  movel([-0.151447, -0.828061, -2.797798, -1.086530, 1.570796, 1.419350],accel_mss,speed_ms,0,blend_radius_m)
  movel([-0.155435, -0.836303, -2.796291, -1.079795, 1.570796, 1.415362],accel_mss,speed_ms,0,blend_radius_m)
  movel([-0.157149, -0.840333, -2.795540, -1.076516, 1.570796, 1.413648],accel_mss,speed_ms,0,blend_radius_m)
  movel([-0.159989, -0.848193, -2.794051, -1.070145, 1.570796, 1.410807],accel_mss,speed_ms,0,blend_radius_m)
  movel([-0.161109, -0.852028, -2.793312, -1.067049, 1.570796, 1.409688],accel_mss,speed_ms,0,blend_radius_m)
  movel([-0.162732, -0.859501, -2.791847, -1.061041, 1.570796, 1.408064],accel_mss,speed_ms,0,blend_radius_m)
  movel([-0.163230, -0.863145, -2.791122, -1.058122, 1.570796, 1.407566],accel_mss,speed_ms,0,blend_radius_m)
  movel([-0.163513, -0.866720, -2.790402, -1.055267, 1.570796, 1.407283],accel_mss,speed_ms,0,blend_radius_m)
  movel([-0.163602, -0.871655, -2.789397, -1.051337, 1.570796, 1.407194],accel_mss,speed_ms,0,blend_radius_m)
  movel([-0.163380, -0.876401, -2.788417, -1.047571, 1.570796, 1.407417],accel_mss,speed_ms,0,blend_radius_m)
  movel([-0.162870, -0.880943, -2.787467, -1.043979, 1.570796, 1.407926],accel_mss,speed_ms,0,blend_radius_m)
  movel([-0.162104, -0.885286, -2.786547, -1.040556, 1.570796, 1.408692],accel_mss,speed_ms,0,blend_radius_m)
  movel([-0.161097, -0.889404, -2.785664, -1.037321, 1.570796, 1.409700],accel_mss,speed_ms,0,blend_radius_m)
  movel([-0.159870, -0.893285, -2.784823, -1.034282, 1.570796, 1.410927],accel_mss,speed_ms,0,blend_radius_m)
  movel([-0.158448, -0.896924, -2.784025, -1.031439, 1.570796, 1.412348],accel_mss,speed_ms,0,blend_radius_m)
  movel([-0.156848, -0.900304, -2.783277, -1.028807, 1.570796, 1.413948],accel_mss,speed_ms,0,blend_radius_m)
  movel([-0.149158, -0.912135, -2.780604, -1.019650, 1.570796, 1.421638],accel_mss,speed_ms,0,blend_radius_m)
  movel([-0.143209, -0.921779, -2.778359, -1.012250, 1.570796, 1.427587],accel_mss,speed_ms,0,blend_radius_m)
  movel([-0.142775, -0.922813, -2.778115, -1.011461, 1.570796, 1.428021],accel_mss,speed_ms,0,blend_radius_m)
  movel([-0.135600, -0.913354, -2.780324, -1.018712, 1.570796, 1.435197],accel_mss,speed_ms,0,blend_radius_m)
  movel([-0.127938, -0.904013, -2.782449, -1.025928, 1.570796, 1.442859],accel_mss,speed_ms,0,blend_radius_m)
  movel([-0.119839, -0.894825, -2.784486, -1.033078, 1.570796, 1.450957],accel_mss,speed_ms,0,blend_radius_m)
  movel([-0.111369, -0.885835, -2.786430, -1.040124, 1.570796, 1.459427],accel_mss,speed_ms,0,blend_radius_m)
  movel([-0.102591, -0.877095, -2.788273, -1.047021, 1.570796, 1.468205],accel_mss,speed_ms,0,blend_radius_m)
  movel([-0.093574, -0.868644, -2.790012, -1.053733, 1.570796, 1.477222],accel_mss,speed_ms,0,blend_radius_m)
  movel([-0.084386, -0.860539, -2.791641, -1.060208, 1.570796, 1.486410],accel_mss,speed_ms,0,blend_radius_m)
  movel([-0.075105, -0.852829, -2.793156, -1.066404, 1.570796, 1.495692],accel_mss,speed_ms,0,blend_radius_m)
  movel([-0.070692, -0.849394, -2.793820, -1.069175, 1.570796, 1.500104],accel_mss,speed_ms,0,blend_radius_m)
  movel([-0.066171, -0.846121, -2.794447, -1.071821, 1.570796, 1.504626],accel_mss,speed_ms,0,blend_radius_m)
  movel([-0.061579, -0.843047, -2.795030, -1.074312, 1.570796, 1.509218],accel_mss,speed_ms,0,blend_radius_m)
  movel([-0.056967, -0.840218, -2.795562, -1.076609, 1.570796, 1.513830],accel_mss,speed_ms,0,blend_radius_m)
  movel([-0.052375, -0.837673, -2.796037, -1.078679, 1.570796, 1.518421],accel_mss,speed_ms,0,blend_radius_m)
  movel([-0.047846, -0.835454, -2.796448, -1.080487, 1.570796, 1.522951],accel_mss,speed_ms,0,blend_radius_m)
  movel([-0.043425, -0.833599, -2.796789, -1.082000, 1.570796, 1.527371],accel_mss,speed_ms,0,blend_radius_m)
  movel([-0.039161, -0.832150, -2.797055, -1.083184, 1.570796, 1.531636],accel_mss,speed_ms,0,blend_radius_m)
  movel([-0.035094, -0.831147, -2.797238, -1.084004, 1.570796, 1.535702],accel_mss,speed_ms,0,blend_radius_m)
  movel([-0.031268, -0.830626, -2.797333, -1.084430, 1.570796, 1.539528],accel_mss,speed_ms,0,blend_radius_m)
  movel([-0.027734, -0.830629, -2.797332, -1.084428, 1.570796, 1.543062],accel_mss,speed_ms,0,blend_radius_m)
  movel([-0.024533, -0.831189, -2.797230, -1.083970, 1.570796, 1.546264],accel_mss,speed_ms,0,blend_radius_m)
  movel([-0.021709, -0.832340, -2.797020, -1.083029, 1.570796, 1.549087],accel_mss,speed_ms,0,blend_radius_m)
  movel([-0.019297, -0.834113, -2.796695, -1.081581, 1.570796, 1.551499],accel_mss,speed_ms,0,blend_radius_m)
  movel([-0.017345, -0.836537, -2.796247, -1.079604, 1.570796, 1.553452],accel_mss,speed_ms,0,blend_radius_m)
  movel([-0.015891, -0.839644, -2.795669, -1.077075, 1.570796, 1.554905],accel_mss,speed_ms,0,blend_radius_m)
  movel([-0.014708, -0.844472, -2.794760, -1.073157, 1.570796, 1.556088],accel_mss,speed_ms,0,blend_radius_m)
  movel([-0.014174, -0.849958, -2.793712, -1.068720, 1.570796, 1.556622],accel_mss,speed_ms,0,blend_radius_m)
  movel([-0.014196, -0.855947, -2.792548, -1.063895, 1.570796, 1.556600],accel_mss,speed_ms,0,blend_radius_m)
  movel([-0.014673, -0.862293, -2.791292, -1.058804, 1.570796, 1.556123],accel_mss,speed_ms,0,blend_radius_m)
  movel([-0.015515, -0.868851, -2.789970, -1.053568, 1.570796, 1.555282],accel_mss,speed_ms,0,blend_radius_m)
  movel([-0.016634, -0.875486, -2.788607, -1.048296, 1.570796, 1.554162],accel_mss,speed_ms,0,blend_radius_m)
  movel([-0.019330, -0.888444, -2.785871, -1.038074, 1.570796, 1.551466],accel_mss,speed_ms,0,blend_radius_m)
  movel([-0.021385, -0.896660, -2.784083, -1.031646, 1.570796, 1.549411],accel_mss,speed_ms,0,blend_radius_m)
  movel([-0.023782, -0.904827, -2.782265, -1.025296, 1.570796, 1.547015],accel_mss,speed_ms,0,blend_radius_m)
  movel([-0.026474, -0.912947, -2.780417, -1.019025, 1.570796, 1.544323],accel_mss,speed_ms,0,blend_radius_m)
  movel([-0.029419, -0.921037, -2.778534, -1.012818, 1.570796, 1.541377],accel_mss,speed_ms,0,blend_radius_m)
  movel([-0.032573, -0.929096, -2.776617, -1.006676, 1.570796, 1.538223],accel_mss,speed_ms,0,blend_radius_m)
  movel([-0.035892, -0.937137, -2.774661, -1.000590, 1.570796, 1.534904],accel_mss,speed_ms,0,blend_radius_m)
  movel([-0.042880, -0.953213, -2.770623, -0.988553, 1.570796, 1.527916],accel_mss,speed_ms,0,blend_radius_m)
  movel([-0.036325, -0.953508, -2.770548, -0.988333, 1.570796, 1.534471],accel_mss,speed_ms,0,blend_radius_m)
  movel([-0.032953, -0.953917, -2.770442, -0.988029, 1.570796, 1.537843],accel_mss,speed_ms,0,blend_radius_m)
  movel([-0.030089, -0.954829, -2.770208, -0.987352, 1.570796, 1.540707],accel_mss,speed_ms,0,blend_radius_m)
  movel([-0.028984, -0.955552, -2.770021, -0.986816, 1.570796, 1.541813],accel_mss,speed_ms,0,blend_radius_m)
  movel([-0.028168, -0.956495, -2.769777, -0.986117, 1.570796, 1.542628],accel_mss,speed_ms,0,blend_radius_m)
  movel([-0.027690, -0.957681, -2.769470, -0.985239, 1.570796, 1.543106],accel_mss,speed_ms,0,blend_radius_m)
  movel([-0.027603, -0.959140, -2.769090, -0.984159, 1.570796, 1.543193],accel_mss,speed_ms,0,blend_radius_m)
  movel([-0.027958, -0.960895, -2.768632, -0.982862, 1.570796, 1.542838],accel_mss,speed_ms,0,blend_radius_m)
  movel([-0.028810, -0.962986, -2.768083, -0.981321, 1.570796, 1.541986],accel_mss,speed_ms,0,blend_radius_m)
  movel([-0.030204, -0.965433, -2.767436, -0.979520, 1.570796, 1.540592],accel_mss,speed_ms,0,blend_radius_m)
  movel([-0.032189, -0.968258, -2.766684, -0.977447, 1.570796, 1.538607],accel_mss,speed_ms,0,blend_radius_m)
  movel([-0.034030, -0.970557, -2.766069, -0.975764, 1.570796, 1.536766],accel_mss,speed_ms,0,blend_radius_m)
  movel([-0.035882, -0.972625, -2.765511, -0.974253, 1.570796, 1.534914],accel_mss,speed_ms,0,blend_radius_m)
  movel([-0.037742, -0.974479, -2.765009, -0.972901, 1.570796, 1.533055],accel_mss,speed_ms,0,blend_radius_m)
  movel([-0.041487, -0.977625, -2.764152, -0.970612, 1.570796, 1.529310],accel_mss,speed_ms,0,blend_radius_m)
  movel([-0.043369, -0.978954, -2.763787, -0.969648, 1.570796, 1.527427],accel_mss,speed_ms,0,blend_radius_m)
  movel([-0.047159, -0.981220, -2.763163, -0.968006, 1.570796, 1.523638],accel_mss,speed_ms,0,blend_radius_m)
  movel([-0.050963, -0.983074, -2.762650, -0.966665, 1.570796, 1.519833],accel_mss,speed_ms,0,blend_radius_m)
  movel([-0.054779, -0.984659, -2.762209, -0.965521, 1.570796, 1.516017],accel_mss,speed_ms,0,blend_radius_m)
  movel([-0.062394, -0.987558, -2.761398, -0.963434, 1.570796, 1.508402],accel_mss,speed_ms,0,blend_radius_m)
  movel([-0.066370, -0.993967, -2.759582, -0.958840, 1.570796, 1.504426],accel_mss,speed_ms,0,blend_radius_m)
  movel([-0.068546, -0.997167, -2.758665, -0.956558, 1.570796, 1.502250],accel_mss,speed_ms,0,blend_radius_m)
  movel([-0.070857, -1.000276, -2.757766, -0.954347, 1.570796, 1.499939],accel_mss,speed_ms,0,blend_radius_m)
  movel([-0.073309, -1.003227, -2.756906, -0.952256, 1.570796, 1.497488],accel_mss,speed_ms,0,blend_radius_m)
  movel([-0.075903, -1.005952, -2.756106, -0.950331, 1.570796, 1.494894],accel_mss,speed_ms,0,blend_radius_m)
  movel([-0.078648, -1.008386, -2.755387, -0.948616, 1.570796, 1.492149],accel_mss,speed_ms,0,blend_radius_m)
  movel([-0.081555, -1.010470, -2.754767, -0.947152, 1.570796, 1.489241],accel_mss,speed_ms,0,blend_radius_m)
  movel([-0.083598, -1.011520, -2.754454, -0.946415, 1.570796, 1.487198],accel_mss,speed_ms,0,blend_radius_m)
  movel([-0.085214, -1.011878, -2.754347, -0.946164, 1.570796, 1.485582],accel_mss,speed_ms,0,blend_radius_m)
  movel([-0.086450, -1.011645, -2.754417, -0.946328, 1.570796, 1.484347],accel_mss,speed_ms,0,blend_radius_m)
  movel([-0.087346, -1.010917, -2.754634, -0.946838, 1.570796, 1.483451],accel_mss,speed_ms,0,blend_radius_m)
  movel([-0.087946, -1.009791, -2.754969, -0.947628, 1.570796, 1.482851],accel_mss,speed_ms,0,blend_radius_m)
  movel([-0.088287, -1.008371, -2.755391, -0.948627, 1.570796, 1.482509],accel_mss,speed_ms,0,blend_radius_m)
  movel([-0.088418, -1.006753, -2.755870, -0.949766, 1.570796, 1.482378],accel_mss,speed_ms,0,blend_radius_m)
  movel([-0.088369, -1.005030, -2.756377, -0.950982, 1.570796, 1.482428],accel_mss,speed_ms,0,blend_radius_m)
  movel([-0.087893, -1.001208, -2.757495, -0.953686, 1.570796, 1.482904],accel_mss,speed_ms,0,blend_radius_m)
  movel([-0.087059, -0.997250, -2.758641, -0.956499, 1.570796, 1.483737],accel_mss,speed_ms,0,blend_radius_m)
  movel([-0.084858, -0.988993, -2.760994, -0.962402, 1.570796, 1.485939],accel_mss,speed_ms,0,blend_radius_m)
  movel([-0.093540, -0.987568, -2.761395, -0.963426, 1.570796, 1.477256],accel_mss,speed_ms,0,blend_radius_m)
  movel([-0.102455, -0.986524, -2.761688, -0.964178, 1.570796, 1.468341],accel_mss,speed_ms,0,blend_radius_m)
  movel([-0.111365, -0.985448, -2.761989, -0.964952, 1.570796, 1.459431],accel_mss,speed_ms,0,blend_radius_m)
  movel([-0.115747, -0.984770, -2.762178, -0.965441, 1.570796, 1.455049],accel_mss,speed_ms,0,blend_radius_m)
  movel([-0.120046, -0.983927, -2.762413, -0.966049, 1.570796, 1.450750],accel_mss,speed_ms,0,blend_radius_m)
  movel([-0.124039, -0.982910, -2.762695, -0.966783, 1.570796, 1.446757],accel_mss,speed_ms,0,blend_radius_m)
  movel([-0.127889, -0.981713, -2.763027, -0.967649, 1.570796, 1.442907],accel_mss,speed_ms,0,blend_radius_m)
  movel([-0.135327, -0.978974, -2.763782, -0.969633, 1.570796, 1.435469],accel_mss,speed_ms,0,blend_radius_m)
  movel([-0.142709, -0.976168, -2.764550, -0.971671, 1.570796, 1.428087],accel_mss,speed_ms,0,blend_radius_m)
  movel([-0.150371, -0.973750, -2.765207, -0.973432, 1.570796, 1.420425],accel_mss,speed_ms,0,blend_radius_m)
  movel([-0.152086, -0.978530, -2.763904, -0.969955, 1.570796, 1.418710],accel_mss,speed_ms,0,blend_radius_m)
  movel([-0.153549, -0.983185, -2.762619, -0.966585, 1.570796, 1.417247],accel_mss,speed_ms,0,blend_radius_m)
  movel([-0.154762, -0.987705, -2.761356, -0.963328, 1.570796, 1.416035],accel_mss,speed_ms,0,blend_radius_m)
  movel([-0.155729, -0.992084, -2.760119, -0.960186, 1.570796, 1.415067],accel_mss,speed_ms,0,blend_radius_m)
  movel([-0.156451, -0.996319, -2.758909, -0.957161, 1.570796, 1.414345],accel_mss,speed_ms,0,blend_radius_m)
  movel([-0.156938, -1.000405, -2.757728, -0.954256, 1.570796, 1.413859],accel_mss,speed_ms,0,blend_radius_m)
  movel([-0.157185, -1.004336, -2.756581, -0.951472, 1.570796, 1.413612],accel_mss,speed_ms,0,blend_radius_m)
  movel([-0.157205, -1.008112, -2.755468, -0.948809, 1.570796, 1.413592],accel_mss,speed_ms,0,blend_radius_m)
  movel([-0.156995, -1.011726, -2.754393, -0.946271, 1.570796, 1.413802],accel_mss,speed_ms,0,blend_radius_m)
  movel([-0.156554, -1.015168, -2.753359, -0.943862, 1.570796, 1.414242],accel_mss,speed_ms,0,blend_radius_m)
  movel([-0.155895, -1.018445, -2.752366, -0.941578, 1.570796, 1.414901],accel_mss,speed_ms,0,blend_radius_m)
  movel([-0.155018, -1.021546, -2.751419, -0.939423, 1.570796, 1.415778],accel_mss,speed_ms,0,blend_radius_m)
  movel([-0.153919, -1.024464, -2.750522, -0.937404, 1.570796, 1.416877],accel_mss,speed_ms,0,blend_radius_m)
  movel([-0.152607, -1.027203, -2.749673, -0.935513, 1.570796, 1.418189],accel_mss,speed_ms,0,blend_radius_m)
  movel([-0.151084, -1.029753, -2.748877, -0.933759, 1.570796, 1.419713],accel_mss,speed_ms,0,blend_radius_m)
  movel([-0.149346, -1.032112, -2.748136, -0.932140, 1.570796, 1.421450],accel_mss,speed_ms,0,blend_radius_m)
  movel([-0.146282, -1.035378, -2.747104, -0.929908, 1.570796, 1.424514],accel_mss,speed_ms,0,blend_radius_m)
  movel([-0.142850, -1.038167, -2.746215, -0.928007, 1.570796, 1.427946],accel_mss,speed_ms,0,blend_radius_m)
  movel([-0.139097, -1.040532, -2.745456, -0.926400, 1.570796, 1.431699],accel_mss,speed_ms,0,blend_radius_m)
  movel([-0.135055, -1.042514, -2.744817, -0.925058, 1.570796, 1.435741],accel_mss,speed_ms,0,blend_radius_m)
  movel([-0.130770, -1.044161, -2.744284, -0.923944, 1.570796, 1.440026],accel_mss,speed_ms,0,blend_radius_m)
  movel([-0.126280, -1.045512, -2.743844, -0.923033, 1.570796, 1.444516],accel_mss,speed_ms,0,blend_radius_m)
  movel([-0.121626, -1.046612, -2.743485, -0.922291, 1.570796, 1.449171],accel_mss,speed_ms,0,blend_radius_m)
  movel([-0.116838, -1.047491, -2.743198, -0.921700, 1.570796, 1.453958],accel_mss,speed_ms,0,blend_radius_m)
  movel([-0.106974, -1.048821, -2.742762, -0.920806, 1.570796, 1.463822],accel_mss,speed_ms,0,blend_radius_m)
  movel([-0.096981, -1.049909, -2.742404, -0.920076, 1.570796, 1.473815],accel_mss,speed_ms,0,blend_radius_m)
  movel([-0.089406, -1.051010, -2.742041, -0.919338, 1.570796, 1.481391],accel_mss,speed_ms,0,blend_radius_m)
  movel([-0.086797, -1.051182, -2.741984, -0.919223, 1.570796, 1.484000],accel_mss,speed_ms,0,blend_radius_m)
  movel([-0.082087, -1.051090, -2.742014, -0.919284, 1.570796, 1.488709],accel_mss,speed_ms,0,blend_radius_m)
  movel([-0.081105, -1.051267, -2.741956, -0.919166, 1.570796, 1.489692],accel_mss,speed_ms,0,blend_radius_m)
  movel([-0.080223, -1.051641, -2.741832, -0.918916, 1.570796, 1.490574],accel_mss,speed_ms,0,blend_radius_m)
  movel([-0.079458, -1.052276, -2.741622, -0.918491, 1.570796, 1.491338],accel_mss,speed_ms,0,blend_radius_m)
  movel([-0.078830, -1.053233, -2.741305, -0.917851, 1.570796, 1.491966],accel_mss,speed_ms,0,blend_radius_m)
  movel([-0.078371, -1.054578, -2.740857, -0.916954, 1.570796, 1.492426],accel_mss,speed_ms,0,blend_radius_m)
  movel([-0.078211, -1.056102, -2.740348, -0.915938, 1.570796, 1.492585],accel_mss,speed_ms,0,blend_radius_m)
  movel([-0.078322, -1.057772, -2.739789, -0.914828, 1.570796, 1.492474],accel_mss,speed_ms,0,blend_radius_m)
  movel([-0.078680, -1.059571, -2.739183, -0.913635, 1.570796, 1.492116],accel_mss,speed_ms,0,blend_radius_m)
  movel([-0.079260, -1.061466, -2.738542, -0.912381, 1.570796, 1.491536],accel_mss,speed_ms,0,blend_radius_m)
  movel([-0.080989, -1.065467, -2.737179, -0.909743, 1.570796, 1.489808],accel_mss,speed_ms,0,blend_radius_m)
  movel([-0.082090, -1.067524, -2.736473, -0.908392, 1.570796, 1.488706],accel_mss,speed_ms,0,blend_radius_m)
  movel([-0.084632, -1.071630, -2.735052, -0.905706, 1.570796, 1.486165],accel_mss,speed_ms,0,blend_radius_m)
  movel([-0.087485, -1.075584, -2.733670, -0.903134, 1.570796, 1.483311],accel_mss,speed_ms,0,blend_radius_m)
  movel([-0.090454, -1.079207, -2.732393, -0.900789, 1.570796, 1.480342],accel_mss,speed_ms,0,blend_radius_m)
  movel([-0.093367, -1.082332, -2.731281, -0.898775, 1.570796, 1.477429],accel_mss,speed_ms,0,blend_radius_m)
  movel([-0.097927, -1.086556, -2.729766, -0.896068, 1.570796, 1.472870],accel_mss,speed_ms,0,blend_radius_m)
  movel([-0.100289, -1.088512, -2.729058, -0.894819, 1.570796, 1.470507],accel_mss,speed_ms,0,blend_radius_m)
  movel([-0.102689, -1.090353, -2.728389, -0.893647, 1.570796, 1.468107],accel_mss,speed_ms,0,blend_radius_m)
  movel([-0.107574, -1.093687, -2.727170, -0.891532, 1.570796, 1.463222],accel_mss,speed_ms,0,blend_radius_m)
  movel([-0.112504, -1.096527, -2.726124, -0.889738, 1.570796, 1.458292],accel_mss,speed_ms,0,blend_radius_m)
  movel([-0.117406, -1.098838, -2.725267, -0.888284, 1.570796, 1.453391],accel_mss,speed_ms,0,blend_radius_m)
  movel([-0.122195, -1.100585, -2.724616, -0.887188, 1.570796, 1.448602],accel_mss,speed_ms,0,blend_radius_m)
  movel([-0.124527, -1.101233, -2.724374, -0.886782, 1.570796, 1.446270],accel_mss,speed_ms,0,blend_radius_m)
  movel([-0.129018, -1.102060, -2.724064, -0.886265, 1.570796, 1.441778],accel_mss,speed_ms,0,blend_radius_m)
  movel([-0.131158, -1.102227, -2.724002, -0.886161, 1.570796, 1.439638],accel_mss,speed_ms,0,blend_radius_m)
  movel([-0.133875, -1.102203, -2.724010, -0.886175, 1.570796, 1.436921],accel_mss,speed_ms,0,blend_radius_m)
  movel([-0.136457, -1.101939, -2.724110, -0.886341, 1.570796, 1.434339],accel_mss,speed_ms,0,blend_radius_m)
  movel([-0.138916, -1.101462, -2.724288, -0.886639, 1.570796, 1.431880],accel_mss,speed_ms,0,blend_radius_m)
  movel([-0.141274, -1.100811, -2.724531, -0.887046, 1.570796, 1.429522],accel_mss,speed_ms,0,blend_radius_m)
  movel([-0.145748, -1.099110, -2.725166, -0.888114, 1.570796, 1.425048],accel_mss,speed_ms,0,blend_radius_m)
  movel([-0.150009, -1.097098, -2.725912, -0.889378, 1.570796, 1.420787],accel_mss,speed_ms,0,blend_radius_m)
  movel([-0.155186, -1.094353, -2.726925, -0.891111, 1.570796, 1.415610],accel_mss,speed_ms,0,blend_radius_m)
  movel([-0.160187, -1.091303, -2.728043, -0.893043, 1.570796, 1.410610],accel_mss,speed_ms,0,blend_radius_m)
  movel([-0.164967, -1.087926, -2.729270, -0.895192, 1.570796, 1.405830],accel_mss,speed_ms,0,blend_radius_m)
  movel([-0.169489, -1.084206, -2.730611, -0.897572, 1.570796, 1.401308],accel_mss,speed_ms,0,blend_radius_m)
  movel([-0.173708, -1.080114, -2.732071, -0.900204, 1.570796, 1.397089],accel_mss,speed_ms,0,blend_radius_m)
  movel([-0.177576, -1.075626, -2.733656, -0.903107, 1.570796, 1.393221],accel_mss,speed_ms,0,blend_radius_m)
  movel([-0.181051, -1.070717, -2.735369, -0.906303, 1.570796, 1.389745],accel_mss,speed_ms,0,blend_radius_m)
  movel([-0.184087, -1.065359, -2.737216, -0.909814, 1.570796, 1.386710],accel_mss,speed_ms,0,blend_radius_m)
  movel([-0.186073, -1.061031, -2.738689, -0.912668, 1.570796, 1.384723],accel_mss,speed_ms,0,blend_radius_m)
  movel([-0.187880, -1.056306, -2.740280, -0.915803, 1.570796, 1.382916],accel_mss,speed_ms,0,blend_radius_m)
  movel([-0.189439, -1.051207, -2.741976, -0.919206, 1.570796, 1.381358],accel_mss,speed_ms,0,blend_radius_m)
  movel([-0.190682, -1.045773, -2.743759, -0.922857, 1.570796, 1.380114],accel_mss,speed_ms,0,blend_radius_m)
  movel([-0.191534, -1.040030, -2.745618, -0.926741, 1.570796, 1.379263],accel_mss,speed_ms,0,blend_radius_m)
  movel([-0.191918, -1.034012, -2.747536, -0.930840, 1.570796, 1.378878],accel_mss,speed_ms,0,blend_radius_m)
  movel([-0.191763, -1.027747, -2.749503, -0.935139, 1.570796, 1.379033],accel_mss,speed_ms,0,blend_radius_m)
  movel([-0.191455, -1.024529, -2.750501, -0.937359, 1.570796, 1.379341],accel_mss,speed_ms,0,blend_radius_m)
  movel([-0.190983, -1.021263, -2.751506, -0.939620, 1.570796, 1.379813],accel_mss,speed_ms,0,blend_radius_m)
  movel([-0.189719, -1.014965, -2.753420, -0.944004, 1.570796, 1.381077],accel_mss,speed_ms,0,blend_radius_m)
  movel([-0.188031, -1.008450, -2.755368, -0.948571, 1.570796, 1.382765],accel_mss,speed_ms,0,blend_radius_m)
  movel([-0.185918, -1.001738, -2.757341, -0.953311, 1.570796, 1.384878],accel_mss,speed_ms,0,blend_radius_m)
  movel([-0.183392, -0.994855, -2.759328, -0.958206, 1.570796, 1.387404],accel_mss,speed_ms,0,blend_radius_m)
  movel([-0.180442, -0.987821, -2.761324, -0.963244, 1.570796, 1.390354],accel_mss,speed_ms,0,blend_radius_m)
  movel([-0.177085, -0.980668, -2.763316, -0.968405, 1.570796, 1.393711],accel_mss,speed_ms,0,blend_radius_m)
  movel([-0.173317, -0.973419, -2.765297, -0.973673, 1.570796, 1.397479],accel_mss,speed_ms,0,blend_radius_m)
  movel([-0.169142, -0.966107, -2.767257, -0.979025, 1.570796, 1.401654],accel_mss,speed_ms,0,blend_radius_m)
  movel([-0.177984, -0.958423, -2.769277, -0.984689, 1.570796, 1.392812],accel_mss,speed_ms,0,blend_radius_m)
  movel([-0.182461, -0.954611, -2.770264, -0.987514, 1.570796, 1.388335],accel_mss,speed_ms,0,blend_radius_m)
  movel([-0.186722, -0.950510, -2.771315, -0.990565, 1.570796, 1.384074],accel_mss,speed_ms,0,blend_radius_m)
  movel([-0.189559, -0.947040, -2.772194, -0.993154, 1.570796, 1.381237],accel_mss,speed_ms,0,blend_radius_m)
  movel([-0.191976, -0.943094, -2.773185, -0.996110, 1.570796, 1.378820],accel_mss,speed_ms,0,blend_radius_m)
  movel([-0.193988, -0.938703, -2.774276, -0.999410, 1.570796, 1.376808],accel_mss,speed_ms,0,blend_radius_m)
  movel([-0.195602, -0.933885, -2.775457, -1.003047, 1.570796, 1.375194],accel_mss,speed_ms,0,blend_radius_m)
  movel([-0.196828, -0.928668, -2.776720, -1.007001, 1.570796, 1.373968],accel_mss,speed_ms,0,blend_radius_m)
  movel([-0.197671, -0.923075, -2.778053, -1.011261, 1.570796, 1.373125],accel_mss,speed_ms,0,blend_radius_m)
  movel([-0.198141, -0.917126, -2.779450, -1.015813, 1.570796, 1.372655],accel_mss,speed_ms,0,blend_radius_m)
  movel([-0.198246, -0.910853, -2.780898, -1.020638, 1.570796, 1.372550],accel_mss,speed_ms,0,blend_radius_m)
  movel([-0.197990, -0.904282, -2.782388, -1.025719, 1.570796, 1.372806],accel_mss,speed_ms,0,blend_radius_m)
  movel([-0.197379, -0.897429, -2.783914, -1.031046, 1.570796, 1.373418],accel_mss,speed_ms,0,blend_radius_m)
  movel([-0.196419, -0.890328, -2.785464, -1.036596, 1.570796, 1.374377],accel_mss,speed_ms,0,blend_radius_m)
  movel([-0.195120, -0.883009, -2.787031, -1.042349, 1.570796, 1.375676],accel_mss,speed_ms,0,blend_radius_m)
  movel([-0.193486, -0.875499, -2.788604, -1.048285, 1.570796, 1.377310],accel_mss,speed_ms,0,blend_radius_m)
  movel([-0.191530, -0.867840, -2.790176, -1.054374, 1.570796, 1.379267],accel_mss,speed_ms,0,blend_radius_m)
  movel([-0.189249, -0.860049, -2.791739, -1.060601, 1.570796, 1.381547],accel_mss,speed_ms,0,blend_radius_m)
  movel([-0.186663, -0.852172, -2.793284, -1.066933, 1.570796, 1.384133],accel_mss,speed_ms,0,blend_radius_m)
  movel([-0.181160, -0.837072, -2.796148, -1.079169, 1.570796, 1.389637],accel_mss,speed_ms,0,blend_radius_m)
  movel([-0.178053, -0.829302, -2.797573, -1.085514, 1.570796, 1.392744],accel_mss,speed_ms,0,blend_radius_m)
  movel([-0.174652, -0.821390, -2.798991, -1.092008, 1.570796, 1.396144],accel_mss,speed_ms,0,blend_radius_m)
  movel([-0.170903, -0.813346, -2.800398, -1.098645, 1.570796, 1.399893],accel_mss,speed_ms,0,blend_radius_m)
  movel([-0.166766, -0.805184, -2.801791, -1.105413, 1.570796, 1.404030],accel_mss,speed_ms,0,blend_radius_m)
  movel([-0.162191, -0.796909, -2.803168, -1.112312, 1.570796, 1.408605],accel_mss,speed_ms,0,blend_radius_m)
  movel([-0.157128, -0.788531, -2.804527, -1.119331, 1.570796, 1.413668],accel_mss,speed_ms,0,blend_radius_m)
  movel([-0.150973, -0.779158, -2.806005, -1.127226, 1.570796, 1.419823],accel_mss,speed_ms,0,blend_radius_m)
  movel([-0.144342, -0.769754, -2.807444, -1.135191, 1.570796, 1.426454],accel_mss,speed_ms,0,blend_radius_m)
  movel([-0.137271, -0.760349, -2.808841, -1.143199, 1.570796, 1.433525],accel_mss,speed_ms,0,blend_radius_m)
  movel([-0.129792, -0.750982, -2.810189, -1.151218, 1.570796, 1.441004],accel_mss,speed_ms,0,blend_radius_m)
  movel([-0.121944, -0.741693, -2.811485, -1.159210, 1.570796, 1.448852],accel_mss,speed_ms,0,blend_radius_m)
  movel([-0.113770, -0.732528, -2.812725, -1.167136, 1.570796, 1.457026],accel_mss,speed_ms,0,blend_radius_m)
  movel([-0.105305, -0.723523, -2.813905, -1.174960, 1.570796, 1.465492],accel_mss,speed_ms,0,blend_radius_m)
  movel([-0.096600, -0.714731, -2.815023, -1.182636, 1.570796, 1.474197],accel_mss,speed_ms,0,blend_radius_m)
  movel([-0.087699, -0.706200, -2.816074, -1.190116, 1.570796, 1.483097],accel_mss,speed_ms,0,blend_radius_m)
  movel([-0.078662, -0.697977, -2.817056, -1.197355, 1.570796, 1.492134],accel_mss,speed_ms,0,blend_radius_m)
  movel([-0.069532, -0.690115, -2.817968, -1.204305, 1.570796, 1.501264],accel_mss,speed_ms,0,blend_radius_m)
  movel([-0.060365, -0.682662, -2.818808, -1.210919, 1.570796, 1.510431],accel_mss,speed_ms,0,blend_radius_m)
  movel([-0.051227, -0.675676, -2.819574, -1.217139, 1.570796, 1.519569],accel_mss,speed_ms,0,blend_radius_m)
  movel([-0.042167, -0.669200, -2.820266, -1.222923, 1.570796, 1.528629],accel_mss,speed_ms,0,blend_radius_m)
  movel([-0.033247, -0.663288, -2.820882, -1.228219, 1.570796, 1.537549],accel_mss,speed_ms,0,blend_radius_m)
  movel([-0.024524, -0.657992, -2.821422, -1.232975, 1.570796, 1.546273],accel_mss,speed_ms,0,blend_radius_m)
  movel([-0.015396, -0.652865, -2.821933, -1.237590, 1.570796, 1.555400],accel_mss,speed_ms,0,blend_radius_m)
  movel([-0.006368, -0.648160, -2.822393, -1.241836, 1.570796, 1.564428],accel_mss,speed_ms,0,blend_radius_m)
  movel([0.002483, -0.644013, -2.822791, -1.245585, 1.570796, 1.573279],accel_mss,speed_ms,0,blend_radius_m)
  movel([0.011077, -0.640576, -2.823116, -1.248698, 1.570796, 1.581874],accel_mss,speed_ms,0,blend_radius_m)
  movel([0.020717, -0.637583, -2.823394, -1.251411, 1.570796, 1.591514],accel_mss,speed_ms,0,blend_radius_m)
  movel([0.029958, -0.635659, -2.823572, -1.253158, 1.570796, 1.600754],accel_mss,speed_ms,0,blend_radius_m)
  movel([0.038695, -0.634822, -2.823648, -1.253918, 1.570796, 1.609491],accel_mss,speed_ms,0,blend_radius_m)
  movel([0.046827, -0.635081, -2.823625, -1.253684, 1.570796, 1.617623],accel_mss,speed_ms,0,blend_radius_m)
  movel([0.054267, -0.636430, -2.823501, -1.252458, 1.570796, 1.625063],accel_mss,speed_ms,0,blend_radius_m)
  movel([0.060928, -0.638861, -2.823276, -1.250252, 1.570796, 1.631725],accel_mss,speed_ms,0,blend_radius_m)
  movel([0.066738, -0.642347, -2.822949, -1.247092, 1.570796, 1.637535],accel_mss,speed_ms,0,blend_radius_m)
  movel([0.071630, -0.646863, -2.822519, -1.243008, 1.570796, 1.642427],accel_mss,speed_ms,0,blend_radius_m)
  movel([0.080139, -0.657114, -2.821510, -1.233765, 1.570796, 1.650935],accel_mss,speed_ms,0,blend_radius_m)
  movel([0.083892, -0.662745, -2.820938, -1.228706, 1.570796, 1.654688],accel_mss,speed_ms,0,blend_radius_m)
  movel([0.087126, -0.669095, -2.820277, -1.223017, 1.570796, 1.657922],accel_mss,speed_ms,0,blend_radius_m)
  movel([0.092254, -0.680122, -2.819089, -1.213178, 1.570796, 1.663050],accel_mss,speed_ms,0,blend_radius_m)
  movel([0.095202, -0.685304, -2.818513, -1.208571, 1.570796, 1.665998],accel_mss,speed_ms,0,blend_radius_m)
  movel([0.098521, -0.690038, -2.817977, -1.204374, 1.570796, 1.669318],accel_mss,speed_ms,0,blend_radius_m)
  movel([0.102318, -0.694152, -2.817503, -1.200734, 1.570796, 1.673114],accel_mss,speed_ms,0,blend_radius_m)
  movel([0.106666, -0.697484, -2.817114, -1.197790, 1.570796, 1.677463],accel_mss,speed_ms,0,blend_radius_m)
  movel([0.111676, -0.699868, -2.816833, -1.195688, 1.570796, 1.682472],accel_mss,speed_ms,0,blend_radius_m)
  movel([0.117434, -0.701139, -2.816682, -1.194568, 1.570796, 1.688231],accel_mss,speed_ms,0,blend_radius_m)
  movel([0.120030, -0.701193, -2.816676, -1.194520, 1.570796, 1.690827],accel_mss,speed_ms,0,blend_radius_m)
  movel([0.122938, -0.700651, -2.816740, -1.194998, 1.570796, 1.693735],accel_mss,speed_ms,0,blend_radius_m)
  movel([0.124501, -0.700063, -2.816810, -1.195517, 1.570796, 1.695297],accel_mss,speed_ms,0,blend_radius_m)
  movel([0.126126, -0.699220, -2.816910, -1.196260, 1.570796, 1.696922],accel_mss,speed_ms,0,blend_radius_m)
  movel([0.127815, -0.698083, -2.817044, -1.197262, 1.570796, 1.698611],accel_mss,speed_ms,0,blend_radius_m)
  movel([0.129555, -0.696612, -2.817217, -1.198560, 1.570796, 1.700351],accel_mss,speed_ms,0,blend_radius_m)
  movel([0.131319, -0.694808, -2.817427, -1.200154, 1.570796, 1.702115],accel_mss,speed_ms,0,blend_radius_m)
  movel([0.132980, -0.692806, -2.817659, -1.201924, 1.570796, 1.703776],accel_mss,speed_ms,0,blend_radius_m)
  movel([0.135970, -0.688482, -2.818155, -1.205753, 1.570796, 1.706767],accel_mss,speed_ms,0,blend_radius_m)
  movel([0.137783, -0.685397, -2.818503, -1.208489, 1.570796, 1.708580],accel_mss,speed_ms,0,blend_radius_m)
  movel([0.139361, -0.682351, -2.818843, -1.211195, 1.570796, 1.710157],accel_mss,speed_ms,0,blend_radius_m)
  movel([0.141870, -0.676394, -2.819497, -1.216498, 1.570796, 1.712666],accel_mss,speed_ms,0,blend_radius_m)
  movel([0.143598, -0.670666, -2.820111, -1.221612, 1.570796, 1.714394],accel_mss,speed_ms,0,blend_radius_m)
  movel([0.144658, -0.665202, -2.820684, -1.226503, 1.570796, 1.715454],accel_mss,speed_ms,0,blend_radius_m)
  movel([0.145152, -0.660066, -2.821212, -1.231111, 1.570796, 1.715948],accel_mss,speed_ms,0,blend_radius_m)
  movel([0.145192, -0.655298, -2.821692, -1.235399, 1.570796, 1.715988],accel_mss,speed_ms,0,blend_radius_m)
  movel([0.144887, -0.650947, -2.822122, -1.239320, 1.570796, 1.715683],accel_mss,speed_ms,0,blend_radius_m)
  movel([0.143440, -0.642970, -2.822890, -1.246529, 1.570796, 1.714237],accel_mss,speed_ms,0,blend_radius_m)
  movel([0.142144, -0.639259, -2.823239, -1.249891, 1.570796, 1.712941],accel_mss,speed_ms,0,blend_radius_m)
  movel([0.140471, -0.635944, -2.823546, -1.252900, 1.570796, 1.711267],accel_mss,speed_ms,0,blend_radius_m)
  movel([0.138417, -0.633061, -2.823809, -1.255519, 1.570796, 1.709214],accel_mss,speed_ms,0,blend_radius_m)
  movel([0.135985, -0.630625, -2.824029, -1.257735, 1.570796, 1.706781],accel_mss,speed_ms,0,blend_radius_m)
  movel([0.133177, -0.628667, -2.824204, -1.259518, 1.570796, 1.703974],accel_mss,speed_ms,0,blend_radius_m)
  movel([0.130010, -0.627194, -2.824334, -1.260860, 1.570796, 1.700806],accel_mss,speed_ms,0,blend_radius_m)
  movel([0.126480, -0.626234, -2.824419, -1.261736, 1.570796, 1.697276],accel_mss,speed_ms,0,blend_radius_m)
  speed_ms = 0.005
  movel([0.126480, -0.620060, -2.817627, -1.274702, 1.570796, 1.697276],accel_mss,speed_ms,0,blend_radius_m)
  speed_ms = 0.040
  movel([0.123325, -0.658068, -2.814003, -1.240318, 1.570796, 1.694121],accel_mss,speed_ms,0,blend_radius_m)
  speed_ms = 0.005
  movel([0.123325, -0.664849, -2.820721, -1.226819, 1.570796, 1.694121],accel_mss,speed_ms,0,blend_radius_m)
  speed_ms = 0.025
  movel([0.118895, -0.664088, -2.820800, -1.227501, 1.570796, 1.689691],accel_mss,speed_ms,0,blend_radius_m)
  movel([0.113905, -0.664232, -2.820785, -1.227372, 1.570796, 1.684701],accel_mss,speed_ms,0,blend_radius_m)
  movel([0.111148, -0.664835, -2.820722, -1.226832, 1.570796, 1.681944],accel_mss,speed_ms,0,blend_radius_m)
  movel([0.108196, -0.665889, -2.820613, -1.225887, 1.570796, 1.678993],accel_mss,speed_ms,0,blend_radius_m)
  movel([0.105036, -0.667465, -2.820448, -1.224476, 1.570796, 1.675833],accel_mss,speed_ms,0,blend_radius_m)
  movel([0.101649, -0.669630, -2.820221, -1.222538, 1.570796, 1.672446],accel_mss,speed_ms,0,blend_radius_m)
  speed_ms = 0.005
  movel([0.101649, -0.662777, -2.813513, -1.236100, 1.570796, 1.672446],accel_mss,speed_ms,0,blend_radius_m)
  speed_ms = 0.040
  movel([0.112275, -0.647453, -2.815075, -1.249862, 1.570796, 1.683072],accel_mss,speed_ms,0,blend_radius_m)
  speed_ms = 0.005
  movel([0.112275, -0.654069, -2.821814, -1.236506, 1.570796, 1.683072],accel_mss,speed_ms,0,blend_radius_m)
  speed_ms = 0.025
  movel([0.112399, -0.649135, -2.822299, -1.240955, 1.570796, 1.683195],accel_mss,speed_ms,0,blend_radius_m)
  movel([0.111517, -0.645203, -2.822678, -1.244509, 1.570796, 1.682314],accel_mss,speed_ms,0,blend_radius_m)
  movel([0.109701, -0.642303, -2.822953, -1.247133, 1.570796, 1.680497],accel_mss,speed_ms,0,blend_radius_m)
  movel([0.107011, -0.640498, -2.823123, -1.248768, 1.570796, 1.677807],accel_mss,speed_ms,0,blend_radius_m)
  movel([0.103521, -0.639825, -2.823186, -1.249378, 1.570796, 1.674318],accel_mss,speed_ms,0,blend_radius_m)
  movel([0.099319, -0.640320, -2.823140, -1.248929, 1.570796, 1.670115],accel_mss,speed_ms,0,blend_radius_m)
  movel([0.094491, -0.642004, -2.822981, -1.247403, 1.570796, 1.665287],accel_mss,speed_ms,0,blend_radius_m)
  movel([0.091867, -0.643305, -2.822858, -1.246225, 1.570796, 1.662663],accel_mss,speed_ms,0,blend_radius_m)
  movel([0.089124, -0.644902, -2.822707, -1.244780, 1.570796, 1.659920],accel_mss,speed_ms,0,blend_radius_m)
  speed_ms = 0.005
  movel([0.089124, -0.638429, -2.815949, -1.258011, 1.570796, 1.659920],accel_mss,speed_ms,0,blend_radius_m)
  speed_ms = 0.040
  movel([0.102652, -0.622712, -2.817393, -1.272283, 1.570796, 1.673448],accel_mss,speed_ms,0,blend_radius_m)
  speed_ms = 0.005
  movel([0.102652, -0.628931, -2.824180, -1.259278, 1.570796, 1.673448],accel_mss,speed_ms,0,blend_radius_m)
  speed_ms = 0.025
  movel([0.102279, -0.626839, -2.824366, -1.261184, 1.570796, 1.673075],accel_mss,speed_ms,0,blend_radius_m)
  movel([0.101580, -0.625025, -2.824525, -1.262839, 1.570796, 1.672376],accel_mss,speed_ms,0,blend_radius_m)
  movel([0.099284, -0.622241, -2.824767, -1.265380, 1.570796, 1.670080],accel_mss,speed_ms,0,blend_radius_m)
  movel([0.095934, -0.620600, -2.824909, -1.266881, 1.570796, 1.666730],accel_mss,speed_ms,0,blend_radius_m)
  movel([0.091712, -0.620117, -2.824950, -1.267322, 1.570796, 1.662509],accel_mss,speed_ms,0,blend_radius_m)
  movel([0.086803, -0.620783, -2.824893, -1.266712, 1.570796, 1.657599],accel_mss,speed_ms,0,blend_radius_m)
  movel([0.081418, -0.622580, -2.824738, -1.265071, 1.570796, 1.652214],accel_mss,speed_ms,0,blend_radius_m)
  movel([0.078603, -0.623902, -2.824623, -1.263863, 1.570796, 1.649399],accel_mss,speed_ms,0,blend_radius_m)
  movel([0.072873, -0.627356, -2.824320, -1.260713, 1.570796, 1.643669],accel_mss,speed_ms,0,blend_radius_m)
  movel([0.070007, -0.629480, -2.824131, -1.258778, 1.570796, 1.640803],accel_mss,speed_ms,0,blend_radius_m)
  speed_ms = 0.005
  movel([0.070007, -0.623252, -2.817345, -1.271791, 1.570796, 1.640803],accel_mss,speed_ms,0,blend_radius_m)
  speed_ms = 0.040
  movel([0.089300, -0.603034, -2.819063, -1.290292, 1.570796, 1.660097],accel_mss,speed_ms,0,blend_radius_m)
  speed_ms = 0.005
  movel([0.089300, -0.608923, -2.825884, -1.277582, 1.570796, 1.660097],accel_mss,speed_ms,0,blend_radius_m)
  speed_ms = 0.025
  movel([0.085848, -0.606670, -2.826066, -1.279652, 1.570796, 1.656644],accel_mss,speed_ms,0,blend_radius_m)
  movel([0.081583, -0.605531, -2.826158, -1.280700, 1.570796, 1.652379],accel_mss,speed_ms,0,blend_radius_m)
  movel([0.076593, -0.605570, -2.826155, -1.280664, 1.570796, 1.647389],accel_mss,speed_ms,0,blend_radius_m)
  movel([0.070948, -0.606830, -2.826054, -1.279505, 1.570796, 1.641744],accel_mss,speed_ms,0,blend_radius_m)
  movel([0.064745, -0.609357, -2.825849, -1.277183, 1.570796, 1.635541],accel_mss,speed_ms,0,blend_radius_m)
  movel([0.061464, -0.611102, -2.825706, -1.275581, 1.570796, 1.632260],accel_mss,speed_ms,0,blend_radius_m)
  movel([0.058084, -0.613171, -2.825536, -1.273682, 1.570796, 1.628881],accel_mss,speed_ms,0,blend_radius_m)
  movel([0.054609, -0.615574, -2.825335, -1.271480, 1.570796, 1.625405],accel_mss,speed_ms,0,blend_radius_m)
  movel([0.051053, -0.618310, -2.825104, -1.268975, 1.570796, 1.621849],accel_mss,speed_ms,0,blend_radius_m)
  movel([0.047438, -0.621372, -2.824842, -1.266175, 1.570796, 1.618234],accel_mss,speed_ms,0,blend_radius_m)
  movel([0.043773, -0.624765, -2.824548, -1.263076, 1.570796, 1.614569],accel_mss,speed_ms,0,blend_radius_m)
  speed_ms = 0.005
  movel([0.043773, -0.618614, -2.817753, -1.276021, 1.570796, 1.614569],accel_mss,speed_ms,0,blend_radius_m)
  speed_ms = 0.040
  movel([0.064233, -0.594251, -2.819759, -1.298379, 1.570796, 1.635029],accel_mss,speed_ms,0,blend_radius_m)
  speed_ms = 0.005
  movel([0.064233, -0.599989, -2.826595, -1.285805, 1.570796, 1.635029],accel_mss,speed_ms,0,blend_radius_m)
  speed_ms = 0.025
  movel([0.063094, -0.597450, -2.826792, -1.288148, 1.570796, 1.633890],accel_mss,speed_ms,0,blend_radius_m)
  movel([0.061364, -0.595588, -2.826934, -1.289867, 1.570796, 1.632160],accel_mss,speed_ms,0,blend_radius_m)
  movel([0.059073, -0.594445, -2.827021, -1.290923, 1.570796, 1.629869],accel_mss,speed_ms,0,blend_radius_m)
  movel([0.056266, -0.594054, -2.827050, -1.291284, 1.570796, 1.627062],accel_mss,speed_ms,0,blend_radius_m)
  movel([0.052290, -0.594549, -2.827013, -1.290827, 1.570796, 1.623086],accel_mss,speed_ms,0,blend_radius_m)
  movel([0.047869, -0.595870, -2.826913, -1.289607, 1.570796, 1.618665],accel_mss,speed_ms,0,blend_radius_m)
  movel([0.042312, -0.598187, -2.826735, -1.287467, 1.570796, 1.613109],accel_mss,speed_ms,0,blend_radius_m)
  movel([0.036448, -0.601320, -2.826491, -1.284578, 1.570796, 1.607244],accel_mss,speed_ms,0,blend_radius_m)
  movel([0.030360, -0.605292, -2.826177, -1.280920, 1.570796, 1.601157],accel_mss,speed_ms,0,blend_radius_m)
  movel([0.024131, -0.610136, -2.825785, -1.276467, 1.570796, 1.594927],accel_mss,speed_ms,0,blend_radius_m)
  movel([0.017873, -0.615862, -2.825311, -1.271216, 1.570796, 1.588669],accel_mss,speed_ms,0,blend_radius_m)
  movel([0.014803, -0.619010, -2.825045, -1.268334, 1.570796, 1.585600],accel_mss,speed_ms,0,blend_radius_m)
  movel([0.008947, -0.625742, -2.824462, -1.262184, 1.570796, 1.579743],accel_mss,speed_ms,0,blend_radius_m)
  movel([0.006216, -0.629270, -2.824150, -1.258969, 1.570796, 1.577013],accel_mss,speed_ms,0,blend_radius_m)
  movel([0.003666, -0.632870, -2.823826, -1.255692, 1.570796, 1.574462],accel_mss,speed_ms,0,blend_radius_m)
  movel([0.001318, -0.636522, -2.823493, -1.252375, 1.570796, 1.572114],accel_mss,speed_ms,0,blend_radius_m)
  speed_ms = 0.005
  movel([0.001318, -0.630181, -2.816719, -1.265488, 1.570796, 1.572114],accel_mss,speed_ms,0,blend_radius_m)
  speed_ms = 0.040
  movel([0.022676, -0.597074, -2.819538, -1.295776, 1.570796, 1.593472],accel_mss,speed_ms,0,blend_radius_m)
  speed_ms = 0.005
  movel([0.022676, -0.602861, -2.826370, -1.283158, 1.570796, 1.593472],accel_mss,speed_ms,0,blend_radius_m)
  speed_ms = 0.025
  movel([0.015376, -0.606334, -2.826093, -1.279962, 1.570796, 1.586173],accel_mss,speed_ms,0,blend_radius_m)
  movel([0.007626, -0.610839, -2.825728, -1.275822, 1.570796, 1.578423],accel_mss,speed_ms,0,blend_radius_m)
  movel([-0.000368, -0.616344, -2.825271, -1.270775, 1.570796, 1.570428],accel_mss,speed_ms,0,blend_radius_m)
  movel([-0.004391, -0.619450, -2.825007, -1.267931, 1.570796, 1.566405],accel_mss,speed_ms,0,blend_radius_m)
  movel([-0.008399, -0.622791, -2.824720, -1.264878, 1.570796, 1.562398],accel_mss,speed_ms,0,blend_radius_m)
  movel([-0.012357, -0.626351, -2.824409, -1.261629, 1.570796, 1.558439],accel_mss,speed_ms,0,blend_radius_m)
  movel([-0.016240, -0.630119, -2.824074, -1.258196, 1.570796, 1.554557],accel_mss,speed_ms,0,blend_radius_m)
  movel([-0.020025, -0.634094, -2.823715, -1.254580, 1.570796, 1.550771],accel_mss,speed_ms,0,blend_radius_m)
  movel([-0.023687, -0.638270, -2.823331, -1.250788, 1.570796, 1.547109],accel_mss,speed_ms,0,blend_radius_m)
  movel([-0.027206, -0.642638, -2.822922, -1.246830, 1.570796, 1.543591],accel_mss,speed_ms,0,blend_radius_m)
  movel([-0.030543, -0.647184, -2.822488, -1.242717, 1.570796, 1.540253],accel_mss,speed_ms,0,blend_radius_m)
  movel([-0.033686, -0.651906, -2.822028, -1.238455, 1.570796, 1.537111],accel_mss,speed_ms,0,blend_radius_m)
  movel([-0.036604, -0.656797, -2.821542, -1.234050, 1.570796, 1.534193],accel_mss,speed_ms,0,blend_radius_m)
  speed_ms = 0.005
  movel([-0.036604, -0.650139, -2.814808, -1.247442, 1.570796, 1.534193],accel_mss,speed_ms,0,blend_radius_m)
  speed_ms = 0.040
  movel([-0.022149, -0.617682, -2.817834, -1.276872, 1.570796, 1.548647],accel_mss,speed_ms,0,blend_radius_m)
  speed_ms = 0.005
  movel([-0.022149, -0.623818, -2.824631, -1.263941, 1.570796, 1.548647],accel_mss,speed_ms,0,blend_radius_m)
  speed_ms = 0.025
  movel([-0.025873, -0.625896, -2.824449, -1.262044, 1.570796, 1.544923],accel_mss,speed_ms,0,blend_radius_m)
  movel([-0.029708, -0.628376, -2.824230, -1.259784, 1.570796, 1.541089],accel_mss,speed_ms,0,blend_radius_m)
  movel([-0.033605, -0.631229, -2.823974, -1.257185, 1.570796, 1.537191],accel_mss,speed_ms,0,blend_radius_m)
  movel([-0.037532, -0.634415, -2.823686, -1.254288, 1.570796, 1.533264],accel_mss,speed_ms,0,blend_radius_m)
  movel([-0.041453, -0.637907, -2.823365, -1.251118, 1.570796, 1.529343],accel_mss,speed_ms,0,blend_radius_m)
  movel([-0.045324, -0.641666, -2.823013, -1.247710, 1.570796, 1.525473],accel_mss,speed_ms,0,blend_radius_m)
  movel([-0.049105, -0.645651, -2.822635, -1.244103, 1.570796, 1.521691],accel_mss,speed_ms,0,blend_radius_m)
  movel([-0.052772, -0.649841, -2.822230, -1.240318, 1.570796, 1.518024],accel_mss,speed_ms,0,blend_radius_m)
  movel([-0.056275, -0.654190, -2.821802, -1.236397, 1.570796, 1.514522],accel_mss,speed_ms,0,blend_radius_m)
  movel([-0.059585, -0.658649, -2.821356, -1.232384, 1.570796, 1.511211],accel_mss,speed_ms,0,blend_radius_m)
  movel([-0.062677, -0.663173, -2.820894, -1.228322, 1.570796, 1.508120],accel_mss,speed_ms,0,blend_radius_m)
  movel([-0.065528, -0.667725, -2.820421, -1.224243, 1.570796, 1.505269],accel_mss,speed_ms,0,blend_radius_m)
  movel([-0.068119, -0.672260, -2.819941, -1.220187, 1.570796, 1.502677],accel_mss,speed_ms,0,blend_radius_m)
  movel([-0.070432, -0.676751, -2.819458, -1.216180, 1.570796, 1.500365],accel_mss,speed_ms,0,blend_radius_m)
  movel([-0.072431, -0.681141, -2.818977, -1.212271, 1.570796, 1.498365],accel_mss,speed_ms,0,blend_radius_m)
  movel([-0.074111, -0.685403, -2.818502, -1.208484, 1.570796, 1.496685],accel_mss,speed_ms,0,blend_radius_m)
  speed_ms = 0.005
  movel([-0.074111, -0.678316, -2.811828, -1.222244, 1.570796, 1.496685],accel_mss,speed_ms,0,blend_radius_m)
  speed_ms = 0.040
  movel([-0.066858, -0.651007, -2.814721, -1.246661, 1.570796, 1.503938],accel_mss,speed_ms,0,blend_radius_m)
  speed_ms = 0.005
  movel([-0.066858, -0.657679, -2.821453, -1.233257, 1.570796, 1.503938],accel_mss,speed_ms,0,blend_radius_m)
  speed_ms = 0.025
  movel([-0.070442, -0.659917, -2.821227, -1.231245, 1.570796, 1.500354],accel_mss,speed_ms,0,blend_radius_m)
  movel([-0.074094, -0.662754, -2.820937, -1.228698, 1.570796, 1.496702],accel_mss,speed_ms,0,blend_radius_m)
  movel([-0.077748, -0.666088, -2.820592, -1.225709, 1.570796, 1.493049],accel_mss,speed_ms,0,blend_radius_m)
  movel([-0.081363, -0.669821, -2.820201, -1.222368, 1.570796, 1.489434],accel_mss,speed_ms,0,blend_radius_m)
  movel([-0.084887, -0.673859, -2.819770, -1.218760, 1.570796, 1.485909],accel_mss,speed_ms,0,blend_radius_m)
  movel([-0.088268, -0.678100, -2.819311, -1.214978, 1.570796, 1.482528],accel_mss,speed_ms,0,blend_radius_m)
  movel([-0.091469, -0.682453, -2.818832, -1.211104, 1.570796, 1.479327],accel_mss,speed_ms,0,blend_radius_m)
  movel([-0.094435, -0.686824, -2.818342, -1.207223, 1.570796, 1.476361],accel_mss,speed_ms,0,blend_radius_m)
  movel([-0.097268, -0.691333, -2.817829, -1.203227, 1.570796, 1.473529],accel_mss,speed_ms,0,blend_radius_m)
  movel([-0.099872, -0.695854, -2.817305, -1.199230, 1.570796, 1.470924],accel_mss,speed_ms,0,blend_radius_m)
  movel([-0.102209, -0.700332, -2.816778, -1.195279, 1.570796, 1.468587],accel_mss,speed_ms,0,blend_radius_m)
  movel([-0.104211, -0.704697, -2.816256, -1.191437, 1.570796, 1.466585],accel_mss,speed_ms,0,blend_radius_m)
  movel([-0.105837, -0.708883, -2.815747, -1.187759, 1.570796, 1.464959],accel_mss,speed_ms,0,blend_radius_m)
  movel([-0.107039, -0.712835, -2.815259, -1.184295, 1.570796, 1.463757],accel_mss,speed_ms,0,blend_radius_m)
  movel([-0.107755, -0.716483, -2.814803, -1.181103, 1.570796, 1.463041],accel_mss,speed_ms,0,blend_radius_m)
  movel([-0.107950, -0.719776, -2.814386, -1.178227, 1.570796, 1.462846],accel_mss,speed_ms,0,blend_radius_m)
  speed_ms = 0.005
  movel([-0.107950, -0.712210, -2.807791, -1.192388, 1.570796, 1.462846],accel_mss,speed_ms,0,blend_radius_m)
  speed_ms = 0.040
  movel([-0.110320, -0.694703, -2.809939, -1.207747, 1.570796, 1.460476],accel_mss,speed_ms,0,blend_radius_m)
  speed_ms = 0.005
  movel([-0.110320, -0.702026, -2.816576, -1.193787, 1.570796, 1.460476],accel_mss,speed_ms,0,blend_radius_m)
  speed_ms = 0.025
  movel([-0.115088, -0.707348, -2.815934, -1.189107, 1.570796, 1.455708],accel_mss,speed_ms,0,blend_radius_m)
  movel([-0.119860, -0.713289, -2.815203, -1.183897, 1.570796, 1.450936],accel_mss,speed_ms,0,blend_radius_m)
  movel([-0.124369, -0.719568, -2.814412, -1.178409, 1.570796, 1.446427],accel_mss,speed_ms,0,blend_radius_m)
  movel([-0.128353, -0.725905, -2.813597, -1.172887, 1.570796, 1.442443],accel_mss,speed_ms,0,blend_radius_m)
  movel([-0.131570, -0.732040, -2.812790, -1.167559, 1.570796, 1.439226],accel_mss,speed_ms,0,blend_radius_m)
  movel([-0.132817, -0.734957, -2.812400, -1.165032, 1.570796, 1.437979],accel_mss,speed_ms,0,blend_radius_m)
  movel([-0.133780, -0.737723, -2.812027, -1.162639, 1.570796, 1.437016],accel_mss,speed_ms,0,blend_radius_m)
  movel([-0.134435, -0.740322, -2.811673, -1.160394, 1.570796, 1.436361],accel_mss,speed_ms,0,blend_radius_m)
  movel([-0.134755, -0.742718, -2.811344, -1.158326, 1.570796, 1.436041],accel_mss,speed_ms,0,blend_radius_m)
  movel([-0.134702, -0.744874, -2.811046, -1.156469, 1.570796, 1.436094],accel_mss,speed_ms,0,blend_radius_m)
  movel([-0.134258, -0.746776, -2.810781, -1.154832, 1.570796, 1.436538],accel_mss,speed_ms,0,blend_radius_m)
  speed_ms = 0.005
  movel([-0.134258, -0.738862, -2.804254, -1.169273, 1.570796, 1.436538],accel_mss,speed_ms,0,blend_radius_m)
  speed_ms = 0.040
  movel([-0.143177, -0.737843, -2.804395, -1.170150, 1.570796, 1.427620],accel_mss,speed_ms,0,blend_radius_m)
  speed_ms = 0.005
  movel([-0.143177, -0.745745, -2.810925, -1.155719, 1.570796, 1.427620],accel_mss,speed_ms,0,blend_radius_m)
  speed_ms = 0.025
  movel([-0.148309, -0.754539, -2.809682, -1.148168, 1.570796, 1.422487],accel_mss,speed_ms,0,blend_radius_m)
  movel([-0.150599, -0.758939, -2.809046, -1.144404, 1.570796, 1.420197],accel_mss,speed_ms,0,blend_radius_m)
  movel([-0.152589, -0.763235, -2.808417, -1.140737, 1.570796, 1.418207],accel_mss,speed_ms,0,blend_radius_m)
  movel([-0.154194, -0.767366, -2.807803, -1.137220, 1.570796, 1.416602],accel_mss,speed_ms,0,blend_radius_m)
  movel([-0.155337, -0.771270, -2.807215, -1.133904, 1.570796, 1.415460],accel_mss,speed_ms,0,blend_radius_m)
  movel([-0.155927, -0.774872, -2.806666, -1.130851, 1.570796, 1.414869],accel_mss,speed_ms,0,blend_radius_m)
  movel([-0.155895, -0.778122, -2.806166, -1.128101, 1.570796, 1.414902],accel_mss,speed_ms,0,blend_radius_m)
  speed_ms = 0.005
  # Splitting Linear movement in 2 (instruction 3386: MoveL 3110)
  movel([-0.155895, -0.758152, -2.790024, -1.164213, 1.570796, 1.414902],accel_mss,speed_ms,0,blend_radius_m)
  movel([-0.155895, -0.740536, -2.773768, -1.198085, 1.570796, 1.414902],accel_mss,speed_ms,0,blend_radius_m)
  speed_ms = 1.000
  movel([-0.155895, -0.740536, -2.773768, -1.198085, 1.570796, 1.414902],accel_mss,speed_ms,0,blend_radius_m)
  # Splitting Linear movement in 6 (instruction 3389: MoveL 3112)
  movel([-0.155895, -0.715708, -2.746447, -1.250234, 1.570796, 1.414902],accel_mss,speed_ms,0,blend_radius_m)
  movel([-0.155895, -0.695699, -2.718871, -1.297819, 1.570796, 1.414902],accel_mss,speed_ms,0,blend_radius_m)
  movel([-0.155895, -0.679715, -2.691064, -1.341610, 1.570796, 1.414902],accel_mss,speed_ms,0,blend_radius_m)
  movel([-0.155895, -0.667122, -2.663045, -1.382222, 1.570796, 1.414902],accel_mss,speed_ms,0,blend_radius_m)
  movel([-0.155895, -0.657412, -2.634827, -1.420150, 1.570796, 1.414902],accel_mss,speed_ms,0,blend_radius_m)
  movel([-0.155895, -0.650173, -2.606417, -1.455798, 1.570796, 1.414902],accel_mss,speed_ms,0,blend_radius_m)
  # End of main program
end

Machining1()
